(* IEC 61131-3 sources: guidance-for-physical-ai-production-designer-on-aws/source/plan2cell/crates/bt2plc/tests/golden/welding_cell_2_small/codesys/head/POU, 2 files *)

(* ---- PLC_PRG.st ---- *)
(*
 * PLC_PRG - Head PLC cell program
 * Generated by bt2plc 0.1.0 for cell welding_cell_2_small (plan bt_1790934549_welding_cell_2_small)
 *
 * Copies every robot's GVL_IO block into the cell's input array, runs FB_Cell and
 * copies the commands back (whole arrays / single bytes only).
 *
 * Operator (plain VARs, pulses are cleared after each scan):
 *   bAutoRun          Level: start a cycle whenever the cell is READY
 *                     (initialised from GVL_Cell.AUTO_RUN on the first scan)
 *   bStart            Pulse: start one cycle
 *   bStop             Pulse: abort (ERR_OPERATOR_STOP); latched in every state, also
 *                     cancels a running reset (CS_RESETTING -> CS_ERROR)
 *   bReset            Pulse: reset after an error (a pulse during CS_ABORTING is kept)
 *   bRecoveryConfirm  Pulse: after an abort mid-cycle or a start-up with an active robot
 *                     away from home, robots moved clear -> sequential blind homing
 *
 * Status: PLC_PRG.fbCell.eState / eError / nErrorRobot / nErrorOp / nErrorZone /
 *         bRecoveryRequired / udiCycles / tLastCycle / aeRobotState / awStep / adwGrant ...
 *
 * Task: MainTask (4 ms cycle)
 *)

PROGRAM PLC_PRG
VAR
    (* Cell controller *)
    fbCell              : FB_Cell;

    (* === Operator === *)
    bAutoRun            : BOOL := TRUE;     (* overwritten by GVL_Cell.AUTO_RUN on the first scan *)
    bStart              : BOOL;
    bStop               : BOOL;
    bReset              : BOOL;
    bRecoveryConfirm    : BOOL;

    (* === Status readback === *)
    eCellState          : E_CellState;
    eCellError          : E_CellError;
    bCellError          : BOOL;
    bRecoveryRequired   : BOOL;
    udiCycles           : UDINT;

    (* Robot input images for fbCell *)
    _astIn              : ARRAY[1..2] OF ST_RobotIn;
    _bFirstScan         : BOOL := TRUE;
END_VAR

(* ---- PLC_PRG_Body.st ---- *)
(*
 * PLC_PRG - Implementation
 *)

IF _bFirstScan THEN
    bAutoRun := GVL_Cell.AUTO_RUN;
    _bFirstScan := FALSE;
END_IF

(* ============================================================================
   INPUTS: GVL_IO -> fbCell (robot -> PLC)
   ============================================================================ *)

(* 1: R1 - robot1 - kuka_robi1 (kuka-robi1, 192.168.100.11) *)
_astIn[1].abySafeIn[0] := GVL_IO.bySafeIn0_R1;
_astIn[1].abySafeIn[1] := GVL_IO.bySafeIn1_R1;
_astIn[1].abySafeIn[2] := GVL_IO.bySafeIn2_R1;
_astIn[1].abySafeIn[3] := GVL_IO.bySafeIn3_R1;
_astIn[1].abySafeIn[4] := GVL_IO.bySafeIn4_R1;
_astIn[1].abySafeIn[5] := GVL_IO.bySafeIn5_R1;
_astIn[1].abySafeIn[6] := GVL_IO.bySafeIn6_R1;
_astIn[1].abySafeIn[7] := GVL_IO.bySafeIn7_R1;
_astIn[1].aVassIn := GVL_IO.aVassInputData_R1;

(* 2: R2 - robot2 - kuka_robi2 (kuka-robi2, 192.168.100.12) *)
_astIn[2].abySafeIn[0] := GVL_IO.bySafeIn0_R2;
_astIn[2].abySafeIn[1] := GVL_IO.bySafeIn1_R2;
_astIn[2].abySafeIn[2] := GVL_IO.bySafeIn2_R2;
_astIn[2].abySafeIn[3] := GVL_IO.bySafeIn3_R2;
_astIn[2].abySafeIn[4] := GVL_IO.bySafeIn4_R2;
_astIn[2].abySafeIn[5] := GVL_IO.bySafeIn5_R2;
_astIn[2].abySafeIn[6] := GVL_IO.bySafeIn6_R2;
_astIn[2].abySafeIn[7] := GVL_IO.bySafeIn7_R2;
_astIn[2].aVassIn := GVL_IO.aVassInputData_R2;

(* ============================================================================
   CELL
   ============================================================================ *)
fbCell(
    bEnable             := TRUE,
    bAutoRun            := bAutoRun,
    bStart              := bStart,
    bStop               := bStop,
    bReset              := bReset,
    bRecoveryConfirm    := bRecoveryConfirm,
    astIn               := _astIn,
    eState              => eCellState,
    eError              => eCellError,
    bError              => bCellError,
    bRecoveryRequired   => bRecoveryRequired,
    udiCycles           => udiCycles);

(* ============================================================================
   OUTPUTS: fbCell -> GVL_IO (PLC -> robot)
   ============================================================================ *)

(* 1: R1 - robot1 *)
GVL_IO.bySafeOut0_R1 := fbCell.astOut[1].abySafeOut[0];
GVL_IO.bySafeOut1_R1 := fbCell.astOut[1].abySafeOut[1];
GVL_IO.bySafeOut2_R1 := fbCell.astOut[1].abySafeOut[2];
GVL_IO.bySafeOut3_R1 := fbCell.astOut[1].abySafeOut[3];
GVL_IO.bySafeOut4_R1 := fbCell.astOut[1].abySafeOut[4];
GVL_IO.bySafeOut5_R1 := fbCell.astOut[1].abySafeOut[5];
GVL_IO.bySafeOut6_R1 := fbCell.astOut[1].abySafeOut[6];
GVL_IO.bySafeOut7_R1 := fbCell.astOut[1].abySafeOut[7];
GVL_IO.aVassOutputData_R1 := fbCell.astOut[1].aVassOut;

(* 2: R2 - robot2 *)
GVL_IO.bySafeOut0_R2 := fbCell.astOut[2].abySafeOut[0];
GVL_IO.bySafeOut1_R2 := fbCell.astOut[2].abySafeOut[1];
GVL_IO.bySafeOut2_R2 := fbCell.astOut[2].abySafeOut[2];
GVL_IO.bySafeOut3_R2 := fbCell.astOut[2].abySafeOut[3];
GVL_IO.bySafeOut4_R2 := fbCell.astOut[2].abySafeOut[4];
GVL_IO.bySafeOut5_R2 := fbCell.astOut[2].abySafeOut[5];
GVL_IO.bySafeOut6_R2 := fbCell.astOut[2].abySafeOut[6];
GVL_IO.bySafeOut7_R2 := fbCell.astOut[2].abySafeOut[7];
GVL_IO.aVassOutputData_R2 := fbCell.astOut[2].aVassOut;

(* One-shot operator buttons *)
bStart := FALSE;
bStop := FALSE;
bReset := FALSE;
bRecoveryConfirm := FALSE;
